(*
    Checks that the library parameter overrides of this test project take
    effect (task 10.1). Expected overrides in the Library Manager:
    CT_CHANNELS 4, CT_BUFFER_LENGTH 1000, AO_WAVEFORM_LENGTH 1000,
    FLOW_BUFFER_LENGTH 100.
*)
FUNCTION_BLOCK FB_ParameterTest EXTENDS TcUnit.FB_TestSuite
VAR
    Ct : MBIDivB.FB_CounterTimer;
    Ao : MBIDivB.FB_AnalogOutput;
END_VAR


OverridesSetArrayBounds();


METHOD PRIVATE OverridesSetArrayBounds

TEST('OverridesSetArrayBounds');

// Element counts from the array sizes (UPPER_BOUND only works on
// variable-length arrays in TwinCAT 3.1.4024).
AssertEquals_UDINT(Expected := 4, Actual := TO_UDINT(SIZEOF(Ct.Channel) / SIZEOF(Ct.Channel[1])), Message := 'CT_CHANNELS');
AssertEquals_UDINT(Expected := 1000, Actual := TO_UDINT(SIZEOF(Ct.Channel[1].Data) / SIZEOF(Ct.Channel[1].Data[1])), Message := 'CT_BUFFER_LENGTH');
AssertEquals_UDINT(Expected := 1000, Actual := TO_UDINT(SIZEOF(Ao.Data) / SIZEOF(Ao.Data[1])), Message := 'AO_WAVEFORM_LENGTH');
AssertEquals_UDINT(Expected := 100, Actual := MBIDivB.GVL_Param.FLOW_BUFFER_LENGTH, Message := 'FLOW_BUFFER_LENGTH');

TEST_FINISHED();
END_METHOD

END_FUNCTION_BLOCK

(* stored: Version 1.1.0.1
   POU FB_ParameterTest: Id {3b6bfc90-2b8a-40c8-b895-d04f2bc2be6a}, SpecialFunc None
   Method OverridesSetArrayBounds: Id {0025bd3e-2822-4acd-8f08-b5280262c6f9} *)
